// TIA Portal V20 export
DATA_BLOCK "HMI_Wartungszähler"   // DB2004
{ S7_Optimized_Access := 'FALSE' }
// stored: AutoNumber false
   VAR RETAIN
      Wartungszähler_Positionierachse_Zyklen : "Wartungszähler_Zyklen";
      Wartungszähler_Positionierachse_Weg { S7_SetPoint := 'True'} : "Wartungszähler_Weg";
      Wartungszähler_Drehachse_Zyklen { S7_SetPoint := 'True'} : "Wartungszähler_Zyklen";
      Wartungszähler_Drehachse_Weg { S7_SetPoint := 'True'} : "Wartungszähler_Weg";
   END_VAR
BEGIN
   Wartungszähler_Positionierachse_Zyklen.Gesamtzyklen := 0;
   Wartungszähler_Positionierachse_Zyklen.Zyklen_soll := 0;
   Wartungszähler_Positionierachse_Zyklen.Zyklen_seit_Wartung := 0;
   Wartungszähler_Positionierachse_Zyklen.Zyklen_bis_Wartung := 500;
   Wartungszähler_Positionierachse_Zyklen.Zähler_reset := FALSE;
   Wartungszähler_Positionierachse_Zyklen.SM_Wartung_fällig := false;
   Wartungszähler_Drehachse_Zyklen.Gesamtzyklen := 0;
   Wartungszähler_Drehachse_Zyklen.Zyklen_soll := 0;
   Wartungszähler_Drehachse_Zyklen.Zyklen_seit_Wartung := 0;
   Wartungszähler_Drehachse_Zyklen.Zyklen_bis_Wartung := 0;
   Wartungszähler_Drehachse_Zyklen.Zähler_reset := FALSE;
   Wartungszähler_Drehachse_Zyklen.SM_Wartung_fällig := false;
END_DATA_BLOCK
